(* CODESYS project 2codesys-pumping-station.project

Project tree, tasks and I/O mapping:
  Device : CODESYS Control Win V3 x64, CODESYS, version 3.5.22.40
    application Application
      libraries: Standard, 3.5.22.0 (System); VisuDialogs, * (System)
      task VISU_TASK (cyclic, interval 100 ms, priority 31) calls VisuElems.Visu_Prg
      task MainTask (cyclic, interval t#20ms, priority 1) calls PLC_PRG
      Enum/
        data type E_StationEtat
        data type E_DefautStation
      Functionblock/
        Station/
          function block FB_Station [ST]
      Function/
        function F_ChangementDePompe [ST]
      program PLC_PRG [ST]
      Structure/
        Station/
          data type ST_StationInput
          data type ST_StationOutput
      visualisation Visualization
      ListeDeTexte/
        text list LT_EtatStation
        text list LT_DefautStation
  libraries: VisuSymbols, 4.5.0.0 (System)
  text list GlobalTextList
*)

// Device/Application/Enum/E_StationEtat
{attribute 'qualified_only'}
{attribute 'strict'}
TYPE E_StationEtat :
(
	Arret, 					// Station arrêtée
	Attente, 				// En attente de la détection du niveau bas
	Demarrage,				// Selection de la pompe
	PompageEnCours,			// Pompage jusqu'à la détection du niveau haut
	Manuel,					// Commande manuelle des pompes par l’opérateur
	Defaut					// Station en état de défaut
);
END_TYPE

// Device/Application/Enum/E_DefautStation
{attribute 'qualified_only'}
{attribute 'strict'}
TYPE E_DefautStation :
(
	Aucun,						// Aucun defaut
	AucunePompeDisponible,		// Les Deux pompes en défaut
	CapteursIncoherents			// Niveau bas et niveau haut TRUE en même temps
);
END_TYPE

// Device/Application/Structure/Station/ST_StationInput
TYPE ST_StationInput :
STRUCT
	xNiveauBas					:	BOOL; // TRUE = niveau bas détecté, démarrage du cycle de pompage demandé
	xNiveauHaut					:	BOOL; // TRUE = niveau haut détecté, arrêt du pompage demandé
	xDemarrageAuto				:	BOOL; // Commande de démarrage automatique de la station
	xArret						:	BOOL; // Commande d'arrêt (TRUE = arrêt demandé)
	xDefautPompe1				:	BOOL; // Retour défaut de la pompe 1
	xDefautPompe2				:	BOOL; // Retour défaut de la pompe 2
	xModeManuel					:	BOOL; // Passage en mode manuel TRUE = manuel, FALSE = automatique
	xDemarragePompe1			:	BOOL; // Demande de démarrage manuel de la pompe 1
	xDemarragePompe2			:	BOOL; // Demande de démarrage manuel de la pompe 2
END_STRUCT
END_TYPE

// Device/Application/Structure/Station/ST_StationOutput
TYPE ST_StationOutput :
STRUCT
	eEtatStation					:	E_StationEtat := E_StationEtat.Arret; 			// Etat actuel de la station
	xPompe1Active					:	BOOL;											// Commande d'activation de la pompe 1
	xPompe2Active					:	BOOL;											// Commande d'activation de la pompe 2
	eDefautStation					:	E_DefautStation := E_DefautStation.Aucun;   	// Catégorie de défaut de la station
	xAlarmePompe1					:	BOOL;											// Signal d'alarme de la pompe 1
	xAlarmePompe2					:	BOOL;											// Signal d'alarme de la pompe 2
	xModeManuelActif				:	BOOL;											// TRUE = mode manuel actif
END_STRUCT						
END_TYPE

// Device/Application/PLC_PRG
PROGRAM PLC_PRG
VAR
	fbStation		:	FB_Station;
	
	xINiveauBas						:	BOOL; 
	xINiveauHaut					:	BOOL; 
	xIDemarrageAuto					:	BOOL; 
	xIArret							:	BOOL; 
	xIDefautPompe1					:	BOOL;
	xIDefautPompe2					:	BOOL;
	xIModeManuel					:	BOOL;
	xIDemarragePompe1				:	BOOL;
	xIDemarragePompe2				:	BOOL;
	
	eOEtatStation					:	E_StationEtat; 			
	xOPompe1Active					:	BOOL;											
	xOPompe2Active					:	BOOL;			
	xOAlarmePompe1					:	BOOL;
	xOAlarmePompe2					:	BOOL;								
	eODefautStation					:	E_DefautStation;   
	xOModeManuelActif				:	BOOL;

	sEtatPompe1						:	WSTRING;
	sEtatPompe2						:	WSTRING;
	xNiveauMoyenAfficher			:	BOOL;
	xNiveauBasAfficher				:	BOOL;
	xNiveauHautAfficher				:	BOOL;
	sModeManuelActifAfficher		:	WSTRING;

END_VAR

fbStation.stInput.xNiveauBas    	:= xINiveauBas;
fbStation.stInput.xNiveauHaut   	:= xINiveauHaut;
fbStation.stInput.xDemarrageAuto	:= xIDemarrageAuto;
fbStation.stInput.xArret        	:= xIArret;
fbStation.stInput.xDefautPompe1 	:= xIDefautPompe1;
fbStation.stInput.xDefautPompe2 	:= xIDefautPompe2;
fbStation.stInput.xModeManuel		:= xIModeManuel;
fbStation.stInput.xDemarragePompe1	:=	xIDemarragePompe1;
fbStation.stInput.xDemarragePompe2	:=	xIDemarragePompe2;


fbStation();


eOEtatStation       := fbStation.stOutput.eEtatStation;
xOPompe1Active      := fbStation.stOutput.xPompe1Active;
xOPompe2Active      := fbStation.stOutput.xPompe2Active;
eODefautStation  	:= fbStation.stOutput.eDefautStation;
xOAlarmePompe1		:= fbStation.stOutput.xAlarmePompe1;
xOAlarmePompe2		:= fbStation.stOutput.xAlarmePompe2;
xOModeManuelActif   := fbStation.stOutput.xModeManuelActif;

xNiveauMoyenAfficher		:=  NOT xINiveauBas AND NOT xINiveauHaut;
xNiveauBasAfficher			:=	xINiveauBas AND NOT xINiveauHaut;
xNiveauHautAfficher			:=	xINiveauHaut AND NOT xINiveauBas;

IF xOPompe1Active THEN
	sEtatPompe1 := "En marche";
ELSIF xOAlarmePompe1 THEN
	sEtatPompe1 := "En Defaut";
ELSE
	sEtatPompe1 := "A l'arrêt";
END_IF

IF xOPompe2Active THEN
	sEtatPompe2 := "En marche";
ELSIF xOAlarmePompe2 THEN
	sEtatPompe2 := "En Defaut";
ELSE
	sEtatPompe2 := "A l'arrêt";
END_IF

IF xOModeManuelActif THEN
	sModeManuelActifAfficher	:=	"oui";
ELSE 
	sModeManuelActifAfficher	:=	"non";
END_IF

END_PROGRAM

// Device/Application/Functionblock/Station/FB_Station
FUNCTION_BLOCK FB_Station

VAR_INPUT
	stInput						:	ST_StationInput;
END_VAR
VAR_OUTPUT
	stOutput					:	ST_StationOutput;
END_VAR
VAR
	iPompePrioritaire			:	INT := 1; // Pompe prioritaire : 1 = pompe 1, 2 = pompe 2
	frontDemarrageAuto			:	R_TRIG; // Front montant du bouton Démarrage auto 
END_VAR

frontDemarrageAuto(CLK 		:= stInput.xDemarrageAuto);
stOutput.xPompe1Active 		:= FALSE;
stOutput.xPompe2Active 		:= FALSE;
stOutput.xAlarmePompe1 		:= stInput.xDefautPompe1;
stOutput.xAlarmePompe2 		:= stInput.xDefautPompe2;


IF NOT stInput.xArret THEN
	// Détection des défauts bloquants (hors arrêt, premier défaut conservé)
	IF stOutput.eEtatStation <> E_StationEtat.Arret
	   AND stOutput.eDefautStation = E_DefautStation.Aucun THEN
		IF stInput.xDefautPompe1 AND stInput.xDefautPompe2 THEN
			stOutput.eDefautStation := E_DefautStation.AucunePompeDisponible;
		ELSIF stInput.xNiveauBas AND stInput.xNiveauHaut THEN
			stOutput.eDefautStation := E_DefautStation.CapteursIncoherents;
		END_IF
	END_IF

	// Un défaut mémorisé force l'état Defaut
	IF stOutput.eDefautStation <> E_DefautStation.Aucun THEN
		stOutput.eEtatStation := E_StationEtat.Defaut;
	END_IF

	CASE stOutput.eEtatStation OF
	//####################################################################################
	E_StationEtat.Arret:
		IF stInput.xModeManuel THEN
			stOutput.eEtatStation := E_StationEtat.Manuel;
		ELSIF frontDemarrageAuto.Q THEN
			stOutput.eEtatStation := E_StationEtat.Attente;
		END_IF
	//####################################################################################	
	E_StationEtat.Attente:
		IF stInput.xNiveauBas THEN
			stOutput.eEtatStation := E_StationEtat.Demarrage;
		END_IF
	//####################################################################################	
	E_StationEtat.Demarrage:
		// Changement de pompe : 
		// Pompe a utiliser en defaut -> lancement de l'autre pompe
		IF stInput.xDefautPompe1 AND (iPompePrioritaire = 1) THEN
			iPompePrioritaire := F_ChangementDePompe(iPompePrioritaire);
		ELSIF stInput.xDefautPompe2 AND (iPompePrioritaire = 2) THEN
			iPompePrioritaire := F_ChangementDePompe(iPompePrioritaire);
		END_IF
		stOutput.eEtatStation := E_StationEtat.PompageEnCours;
	//####################################################################################	
	E_StationEtat.PompageEnCours:
		// Si la pompe prioritaire actuelle tombe en défaut, on bascule sur l'autre
		IF (iPompePrioritaire = 1) AND stInput.xDefautPompe1 THEN
			iPompePrioritaire := 2;
		ELSIF (iPompePrioritaire = 2) AND stInput.xDefautPompe2 THEN
			iPompePrioritaire := 1;
		END_IF
		
		// Pilotage des sorties selon la pompe prioritaire validée
		IF iPompePrioritaire = 1 AND NOT stInput.xDefautPompe1 THEN
			stOutput.xPompe1Active := TRUE;
		ELSIF iPompePrioritaire = 2 AND NOT stInput.xDefautPompe2 THEN
			stOutput.xPompe2Active := TRUE;
		END_IF
				
		// Condition de fin de cycle (Niveau Haut)
		IF stInput.xNiveauHaut THEN
			iPompePrioritaire := F_ChangementDePompe(iPompePrioritaire);
			stOutput.eEtatStation := E_StationEtat.Attente;
		END_IF

	//####################################################################################
	E_StationEtat.Manuel:
		IF NOT stInput.xModeManuel THEN
			stOutput.eEtatStation := E_StationEtat.Arret;
		ELSIF stInput.xDemarragePompe1 AND NOT stInput.xDefautPompe1 THEN
			stOutput.xPompe1Active := TRUE;
		ELSIF stInput.xDemarragePompe2 AND NOT stInput.xDefautPompe2 THEN
			stOutput.xPompe2Active := TRUE;
		END_IF
	//####################################################################################	
	E_StationEtat.Defaut:
		// La Station est en defaut
END_CASE
ELSE 
	stOutput.eDefautStation := E_DefautStation.Aucun;
	stOutput.eEtatStation := E_StationEtat.Arret;
END_IF
stOutput.xModeManuelActif	:= (stOutput.eEtatStation = E_StationEtat.Manuel);

END_FUNCTION_BLOCK

// Device/Application/Function/F_ChangementDePompe
FUNCTION F_ChangementDePompe : INT
VAR_INPUT
	iPompeActuelle		:	INT; // Prend le numero de la pompe actuelle ( 1 ou 2 )
END_VAR
VAR
END_VAR

IF iPompeActuelle = 1 THEN
	F_ChangementDePompe := 2;
ELSIF iPompeActuelle = 2 THEN
	F_ChangementDePompe := 1;
ELSE 
	F_ChangementDePompe := 0;
END_IF

END_FUNCTION

// Device/Application/Visualization
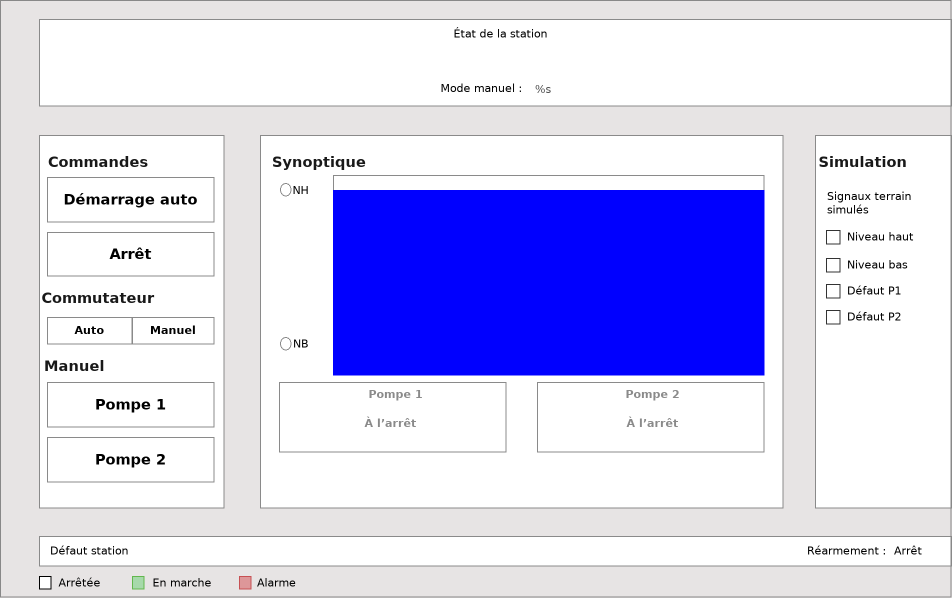
VISUALIZATION Visualization  // 952x598
    RoundedRectangle (39,19 913x87)
    Label (291,0 419x68), "État de la station"
    Label (377,71 230x35), "Mode manuel :"
    RoundedRectangle (39,135 185x373)
    RoundedRectangle (260,135 523x373)
    RoundedRectangle (815,135 137x373)
    RoundedRectangle (39,536 913x30)
    Label (39,144 118x36), "Commandes"
    RoundedRectangle (47,177 167x45), "Démarrage auto", colour toggle: PLC_PRG.xIDemarrageAuto
        tap PLC_PRG.xIDemarrageAuto
    RoundedRectangle (47,232 167x44), "Arrêt", colour toggle: PLC_PRG.xIArret
        OnMouseClick:  ToggleVariable=PLC_PRG.xIArret
    Label (39,280 118x36), "Commutateur"
    RoundedRectangle (47,382 167x45), "Pompe 1", colour toggle: PLC_PRG.xIDemarragePompe1
        OnMouseClick:  ToggleVariable=PLC_PRG.xIDemarragePompe1
    Label (5,348 139x36), "Manuel"
    RoundedRectangle (47,437 167x45), "Pompe 2", colour toggle: PLC_PRG.xIDemarragePompe2
        OnMouseClick:  ToggleVariable=PLC_PRG.xIDemarragePompe2
    RoundedRectangle (47,317 85x27), "Auto", colour toggle: NOT PLC_PRG.xIModeManuel
        OnMouseClick: execute { PLC_PRG.xIModeManuel := FALSE; }
    RoundedRectangle (132,317 82x27), "Manuel", colour toggle: PLC_PRG.xIModeManuel
        OnMouseClick: execute { PLC_PRG.xIModeManuel := TRUE; }
    Line (239,403)
    Label (260,144 118x36), "Synoptique"
    Label (804,144 118x36), "Simulation"
    RoundedRectangle (333,175 431x193)
    RoundedRectangle (279,382 227x70), colour toggle: PLC_PRG.xIDefautPompe1
    RoundedRectangle (537,382 227x70), colour toggle: PLC_PRG.xIDefautPompe2
    Ellipse (280,183 11x13), colour toggle: PLC_PRG.xINiveauHaut
    Ellipse (280,337 11x13), colour toggle: PLC_PRG.xINiveauBas
    Label (279,175 44x31), "NH"
    Label (279,327 44x34), "NB"
    Label (824,175 128x56), "Signaux terrain simulés"
    Checkbox (824,226 122x22), "Niveau haut", variable: PLC_PRG.xINiveauHaut
    Checkbox (824,254 122x22), "Niveau bas", variable: PLC_PRG.xINiveauBas
    Checkbox (824,280 122x22), "Défaut P1", variable: PLC_PRG.xIDefautPompe1
    Checkbox (824,306 122x22), "Défaut P2", variable: PLC_PRG.xIDefautPompe2
    Label (47,536 97x30), "Défaut station :"
    Label (804,536 97x30), "Réarmement :"
    Label (891,536 61x30), "Arrêt"
    Rectangle (39,576 12x13)
    Label (47,568 65x30), "Arrêtée"
    Rectangle (132,576 12x13)
    Label (140,568 84x30), "En marche"
    Rectangle (239,576 12x13)
    Label (244,568 65x30), "Alarme"
    Rectangle (249,47 508x30), text list: 'LT_EtatStation', text index: PLC_PRG.eOEtatStation
    Rectangle (132,542 316x18), text list: 'LT_DefautStation', text index: PLC_PRG.eODefautStation
    Rectangle (338,385 115x19), "Pompe 1", colour toggle: PLC_PRG.xIDefautPompe1
    Rectangle (338,414 115x19), "%s", text variable: PLC_PRG.sEtatPompe1, colour toggle: PLC_PRG.xIDefautPompe1
    Rectangle (595,385 115x19), "Pompe 2", colour toggle: PLC_PRG.xIDefautPompe2
    Rectangle (595,414 115x19), "%s", text variable: PLC_PRG.sEtatPompe2, colour toggle: PLC_PRG.xIDefautPompe2
    RoundedRectangle (333,338 431x30), invisible if: NOT PLC_PRG.xNiveauBasAfficher
    RoundedRectangle (333,264 431x104), invisible if: NOT PLC_PRG.xNiveauMoyenAfficher
    RoundedRectangle (333,190 431x185), invisible if: NOT PLC_PRG.xNiveauHautAfficher
    RoundedRectangle (537,382 227x70), invisible if: PLC_PRG.xOPompe2Active OR PLC_PRG.xIDefautPompe2
    Rectangle (595,385 115x19), "Pompe 2", invisible if: PLC_PRG.xOPompe2Active OR PLC_PRG.xIDefautPompe2
    Rectangle (595,414 115x19), "À l’arrêt", text variable: PLC_PRG.sEtatPompe1, invisible if: PLC_PRG.xOPompe2Active OR PLC_PRG.xIDefautPompe2
    RoundedRectangle (279,382 227x70), invisible if: PLC_PRG.xOPompe1Active OR PLC_PRG.xIDefautPompe1
    Rectangle (338,385 115x19), "Pompe 1", invisible if: PLC_PRG.xOPompe1Active OR PLC_PRG.xIDefautPompe1
    Rectangle (333,414 115x19), "À l’arrêt", text variable: PLC_PRG.sEtatPompe1, invisible if: PLC_PRG.xOPompe1Active OR PLC_PRG.xIDefautPompe1
    Rectangle (532,79 113x21), "%s", text variable: PLC_PRG.sModeManuelActifAfficher
END_VISUALIZATION

(* text list LT_EtatStation (id | default)
  0 | Arrêt
  1 | En attente
  2 | En démarrage
  3 | Pompage en cours
  4 | Mode manuel
  5 | En défaut
   |  *)

(* text list LT_DefautStation (id | default)
  0 | Aucun défaut
  1 | Aucune pompe disponible
  2 | Capteurs incohérents
   |  *)
